Staubli VAL3: updateBtn.pgx

public program updateBtn(num x_nItemIn, string x_sComment)
  local num l_nI
  local num l_nPos
  local string l_sLongStr
  local string l_sBtnText[8]
begin
  switch sLanguage
    case "chinese"
      l_sLongStr=sHmiCN[x_nItemIn]
    break
    //
    case "english"
      l_sLongStr=sHmiEN[x_nItemIn]
    break
  endSwitch
  nBtnItem=x_nItemIn
  //
  for l_nI= 0 to 7
    l_nPos=find(l_sLongStr,",")
    if l_nPos!=-1
      l_sBtnText[l_nI]=left(l_sLongStr,l_nPos)
      l_sLongStr=delete(l_sLongStr,l_nPos+1,0)
    else
      l_sBtnText[l_nI]=l_sLongStr
    endIf
    if l_sBtnText[l_nI]!="Null"
      utBtn_Bottom[l_nI].Common.sText=l_sBtnText[l_nI]
      utBtn_Bottom[l_nI].Appearance.bVisibility=true
    else
      utBtn_Bottom[l_nI].Common.sText=""
      utBtn_Bottom[l_nI].Appearance.bVisibility=false
    endIf
  endFor
end
